(* IEC 61131-3 sources: PortalRobot/Portal_robot/Device/application/ST/ST_HMI, 6 files *)

(* ---- E_HMI_MANUAL_REJECT.st ---- *)
{attribute 'qualified_only'}
{attribute 'strict'}
TYPE E_HMI_MANUAL_REJECT :
(
	NONE,
	HMI_OFFLINE,
	MANUAL_MODE_REQUIRED,
	MODBUS_ACTIVE,
	GLOBAL_ERROR_JOG_ONLY,
	DRIVE_ERROR,
	DRIVES_DISABLED,
	AXIS_BUSY,
	AXIS_NOT_HOMED,
	SOFT_LIMIT,
	COMMAND_CONFLICT,
	ROBOT_BUSY,
	ACTION_ALREADY_REACHED,
	EXTERNAL_ROBOT_NOT_READY,
	MOTION_NOT_READY,
	HATCH_CLOSED,
	CALIBRATION_POINT_UNAVAILABLE
);
END_TYPE

(* ---- ST_AXIS_HMI_COMMAND.st ---- *)
TYPE ST_AXIS_HMI_COMMAND :
STRUCT
	xJogPositive      : BOOL; // Удерживаемый Jog в положительном направлении
	xJogNegative      : BOOL; // Удерживаемый Jog в отрицательном направлении
	{attribute 'symbol' := 'read'}
	xHome             : BOOL; // Импульс поиска домашней позиции выбранной оси
	{attribute 'symbol' := 'read'}
	xMoveAbsolute     : BOOL; // Импульс абсолютного перемещения к lrTargetPosition
	{attribute 'symbol' := 'read'}
	xMoveRelative     : BOOL; // Импульс относительного перемещения на lrRelativeDistance
	lrTargetPosition  : LREAL; // Целевая абсолютная координата оси
	lrRelativeDistance : LREAL; // Подготовленная дистанция относительного движения
END_STRUCT
END_TYPE

(* ---- ST_AXIS_HMI_STATUS.st ---- *)
TYPE ST_AXIS_HMI_STATUS :
STRUCT
	xJogPositiveAllowed   : BOOL; // PLC разрешает положительный Jog
	xJogNegativeAllowed   : BOOL; // PLC разрешает отрицательный Jog
	xHomeAllowed          : BOOL; // PLC разрешает поиск домашней позиции
	xMoveAbsoluteAllowed  : BOOL; // PLC разрешает абсолютное движение
	xMoveRelativePositiveAllowed : BOOL; // PLC разрешает положительный короткий шаг
	xMoveRelativeNegativeAllowed : BOOL; // PLC разрешает отрицательный короткий шаг
	xDriveReady           : BOOL; // Ось включена и готова к движению
	xBusy                 : BOOL; // Ось выполняет ручную команду
	xError                : BOOL; // На оси есть ошибка
	xHomed                : BOOL; // Ось прошла поиск домашней позиции
	lrActualPosition      : LREAL; // Фактическая координата
	lrTargetPosition      : LREAL; // Принятая целевая координата
	lrDeviation           : LREAL; // Отклонение фактической координаты от цели
	lrMinPosition         : LREAL; // Нижний программный предел
	lrMaxPosition         : LREAL; // Верхний программный предел
	lrCommandVelocity     : LREAL; // Фактически заданная скорость ручного движения
	lrMaxVelocity         : LREAL; // Скорость, соответствующая 100 процентам
	eRejectReason         : E_HMI_MANUAL_REJECT; // Числовая причина недоступности команды
	eState                : E_AXIS_STATE; // Числовое состояние автомата оси
END_STRUCT
END_TYPE

(* ---- ST_HMI.st ---- *)
TYPE ST_HMI :
STRUCT
	ActualX : LREAL; // Текущая координата X для существующей визуализации
	ActualY : LREAL; // Текущая координата Y для существующей визуализации
	ActualZ : LREAL; // Текущая координата Z для существующей визуализации
END_STRUCT
END_TYPE

(* ---- ST_PHYSICAL_IO_EVENT.st ---- *)
TYPE ST_PHYSICAL_IO_EVENT :
STRUCT
    udiSequence : UDINT;
    uliTimeMs : ULINT; // Монотонное время от старта приложения, без переполнения TIME
    usiDirection : USINT; // 1 DI; 2 DO
    uiIndex : UINT; // DI 1..84; DO 1..50, index из карты I/O
    usiKind : USINT; // 1 клемма DI; 2 вход программы; 3 DO; 4 подмена DI; 5/6 снять DI; 7 ручной DO; 8/9 возврат DO оператором/программе
    xOld : BOOL;
    xNew : BOOL;
END_STRUCT
END_TYPE

(* ---- ST_ROBOT_HMI_STATUS.st ---- *)
TYPE ST_ROBOT_HMI_STATUS :
STRUCT
	xDrivesPowered       : BOOL; // Все три привода фактически включены
	xDrivesOff           : BOOL; // Все три привода и группа фактически отключены
	xPowerTransitionActive : BOOL; // Выполняется последовательность включения или отключения
	xDrivesEnableAllowed : BOOL; // PLC разрешает включение приводов
	xDrivesDisableAllowed : BOOL; // PLC разрешает отключение приводов
	xResetAllowed        : BOOL; // PLC разрешает команду сброса ручного управления
	xStopAllowed         : BOOL; // PLC разрешает контролируемую остановку
	xPointsAllowed        : BOOL; // PLC разрешает переход к именованной точке
	xGripperAllowed       : BOOL; // PLC разрешает действие захвата
	xGripper1OpenAllowed  : BOOL;
	xGripper1CloseAllowed : BOOL;
	xGripper2OpenAllowed  : BOOL;
	xGripper2CloseAllowed : BOOL;
	xRotateToBlankAllowed : BOOL;
	xRotateToDetailAllowed : BOOL;
	xCommandBusy          : BOOL;
	uiActiveAction        : UINT;
	uiActivePoint         : UINT;
	eRejectReason         : E_HMI_MANUAL_REJECT; // Числовая причина недоступности команды
END_STRUCT
END_TYPE
